{region 'Documentation'}
(*!
<summary>Check equality between consecutive active observations.</summary>
<description>

The first active observation establishes a baseline without deciding a result. Disabling
observation invalidates that baseline, not the held Result. Re-enabling first establishes a new
baseline; Reset clears history.

ObserveFirstCycle FALSE delays the first observation by one enabled call.

</description>
*)
{endregion}
FUNCTION_BLOCK AssertNoValueChange_DT EXTENDS AssertionBase
VAR_INPUT
    IN : DT; //! Actual value to observe.
END_VAR
VAR
    FINPrevious : DT;
    FObservationPrevious : BOOL;
    FEvaluationActive : BOOL;
END_VAR

SUPER^();

{region 'Documentation'}
(*!
<summary>Observe the current value before evaluating a change against the previous observation.</summary>
*)
{endregion}
METHOD PROTECTED Assert
VAR
    PreviousValue : DT;
    Message : STRING(GVL_Constants.MessageLength);
    PreviousText : STRING(GVL_Constants.AssertionValueLength);
    ActualText : STRING(GVL_Constants.AssertionValueLength);
END_VAR
FEvaluationActive := ObservationActive AND FObservationPrevious;
FObservationPrevious := ObservationActive;

IF NOT ObservationActive THEN
    RETURN;
END_IF;

PreviousValue := FINPrevious;
FINPrevious := IN;

IF NOT EvaluationActive THEN
    RETURN;
END_IF;

IF Result = E_Result.Error THEN
    RETURN;
END_IF;

IF Result = E_Result.Failed THEN
    RETURN;
END_IF;

IF IN <> PreviousValue THEN
    PreviousText := DT_TO_STRING(PreviousValue);
    ActualText := DT_TO_STRING(IN);
    Message := CONCAT('Assertion failed: value changed unexpectedly. Previous = ',
        PreviousText);
    Message := CONCAT(Message, ', Actual = ');
    Message := CONCAT(Message, ActualText);
    Message := CONCAT(Message, '.');
    Fail(Message := Message);
    RETURN;
END_IF;

Pass();
END_METHOD

{region 'Documentation'}
(*!
<summary>Current/last call has an active observation and a preceding observation
baseline.</summary>
*)
{endregion}
{attribute 'monitoring' := 'call'}
PROPERTY PUBLIC EvaluationActive : BOOL //! Current/last call has an active observation and a preceding observation baseline.
GET // PUBLIC
EvaluationActive := FEvaluationActive;
END_GET
END_PROPERTY

{region 'Documentation'}
(*!
<summary>Clear observation history and the current evaluation gate.</summary>
*)
{endregion}
METHOD PROTECTED ResetAssertion
FINPrevious := DT#1970-01-01-00:00:00;
FObservationPrevious := FALSE;
FEvaluationActive := FALSE;
END_METHOD

END_FUNCTION_BLOCK

(* stored: Version 1.1.0.1
   POU AssertNoValueChange_DT: Id {f7613b86-0202-4670-a328-890632511b7f}, SpecialFunc None
   Folder Internal: Id {739a2076-50fd-49a9-8518-0a850e0af746}
   Method Assert: Id {557d48b3-26d9-4197-a667-8ea02e1b74f0}
   Property EvaluationActive: Id {f7c85d86-bdcb-462c-8080-0dddae729daa}
   Get Get: Id {a4956aed-c688-4e27-bb7d-af228fe57a79}
   Method ResetAssertion: Id {dcdfaa2d-8838-429d-9c1a-11307000e392} *)
